      [55]
        bool bMarked
        jointRx jJointRx = {j1=119.753729, j2=-7.953574, j3=74.820625, j4=-173.223401, j5=72.415611, j6=-212.309715}
        pointRx pInter
        paraItem pParaItem
          [0]
            bool bSafePoint
            ifItem iIfItem
              [0]
                bool bANDOR[2]
                num nSigIndex[3]
                num nSigType[3]
                num nValue[3]
            mdesc mMdesc = {leave=0}
            num nActionIndex = 41
            num nDelay = 1
            num nMoveType = 1
            num nPercentage
            num nSigValue
        pointRx pPointRx[2] = {x=-39.963894, y=381.881422, z=1281.672322, rx=1.496816, ry=8.299138, rz=89.69815, shoulder=lefty, elbow=epositive, wrist=wpositive}
        string sID
      [56]
        bool bMarked
        jointRx jJointRx = {j1=126.372801, j2=0.947016, j3=58.247522, j4=-173.633502, j5=65.467797, j6=-219.528921}
        pointRx pInter
        paraItem pParaItem
          [0]
            bool bSafePoint
            ifItem iIfItem
              [0]
                bool bANDOR[2]
                num nSigIndex[3]
                num nSigType[3]
                num nValue[3]
            mdesc mMdesc = {leave=0}
            num nActionIndex = 41
            num nDelay = 1
            num nMoveType = 1
            num nPercentage
            num nSigValue
        pointRx pPointRx[2] = {x=-110.0468221, y=381.881454, z=1352.0109929, rx=1.496598, ry=8.298005, rz=89.698483, shoulder=lefty, elbow=epositive, wrist=wpositive}
        string sID
      [57]
        bool bMarked
        jointRx jJointRx = {j1=135.765404, j2=12.255762, j3=45.397511, j4=-174.78792, j5=64.742909, j6=-228.47546}
        pointRx pInter
        paraItem pParaItem
          [0]
            bool bSafePoint
            ifItem iIfItem
              [0]
                bool bANDOR[2]
                num nSigIndex[3]
                num nSigType[3]
                num nValue[3]
            mdesc mMdesc = {leave=0}
            num nActionIndex = 41
            num nDelay = 1
            num nMoveType = 1
            num nPercentage
            num nSigValue
        pointRx pPointRx[2] = {x=-234.761691, y=381.497821, z=1353.29132, rx=1.49622, ry=8.29735, rz=89.698646, shoulder=lefty, elbow=epositive, wrist=wpositive}
        string sID
      [58]
        bool bMarked
        jointRx jJointRx = {j1=138.772753, j2=12.465275, j3=53.540842, j4=-175.467559, j5=73.29136, j6=-230.546088}
        pointRx pInter
        paraItem pParaItem
          [0]
            bool bSafePoint
            ifItem iIfItem
              [0]
                bool bANDOR[2]
                num nSigIndex[3]
                num nSigType[3]
                num nValue[3]
            mdesc mMdesc = {leave=0}
            num nActionIndex = 41
            num nDelay = 1
            num nMoveType = 1
            num nPercentage
            num nSigValue
        pointRx pPointRx[2] = {x=-284.713057, y=381.881445, z=1282.27146, rx=1.496715, ry=8.298986, rz=89.698256, shoulder=lefty, elbow=epositive, wrist=wpositive}
        string sID
      [59]
        bool bMarked
        jointRx jJointRx = {j1=142.602482, j2=20.481815, j3=43.70957, j4=-175.946983, j5=71.740182, j6=-234.319694}
        pointRx pInter
        paraItem pParaItem
          [0]
            bool bSafePoint
            ifItem iIfItem
              [0]
                bool bANDOR[2]
                num nSigIndex[3]
                num nSigType[3]
                num nValue[3]
            mdesc mMdesc = {leave=0}
            num nActionIndex = 41
            num nDelay = 1
            num nMoveType = 1
            num nPercentage
            num nSigValue
        pointRx pPointRx[2] = {x=-357.530662, y=381.881364, z=1278.257011, rx=1.496095, ry=8.297308, rz=89.698645, shoulder=lefty, elbow=epositive, wrist=wpositive}
        string sID
      [60]
        bool bMarked
        jointRx jJointRx = {j1=146.225971, j2=34.147401, j3=22.485673, j4=-176.265369, j5=64.412135, j6=-238.261186}
        pointRx pInter
        paraItem pParaItem
          [0]
            bool bSafePoint
            ifItem iIfItem
              [0]
                bool bANDOR[2]
                num nSigIndex[3]
                num nSigType[3]
                num nValue[3]
            mdesc mMdesc = {leave=0}
            num nActionIndex = 41
            num nDelay = 1
            num nMoveType = 1
            num nPercentage
            num nSigValue
        pointRx pPointRx[2] = {x=-439.57558, y=381.88118, z=1286.715302, rx=1.495603, ry=8.296388, rz=89.698782, shoulder=lefty, elbow=epositive, wrist=wpositive}
        string sID
      [61]
        bool bMarked
        jointRx jJointRx = {j1=145.163516, j2=25.787023, j3=46.647021, j4=-176.436157, j5=80.123032, j6=-236.204112}
        pointRx pInter
        paraItem pParaItem
          [0]
            bool bSafePoint
            ifItem iIfItem
              [0]
                bool bANDOR[2]
                num nSigIndex[3]
                num nSigType[3]
                num nValue[3]
            mdesc mMdesc = {leave=0}
            num nActionIndex = 41
            num nDelay = 1
            num nMoveType = 1
            num nPercentage
            num nSigValue
        pointRx pPointRx[2] = {x=-433.595736, y=395.563274, z=1186.609873, rx=1.496133, ry=8.298356, rz=89.698378, shoulder=lefty, elbow=epositive, wrist=wpositive}
        string sID
      [62]
        bool bMarked
        jointRx jJointRx = {j1=141.740249, j2=16.896756, j3=58.529423, j4=-176.00804128, j5=82.891986, j6=-232.685997}
        pointRx pInter
        paraItem pParaItem
          [0]
            bool bSafePoint
            ifItem iIfItem
              [0]
                bool bANDOR[2]
                num nSigIndex[3]
                num nSigType[3]
                num nValue[3]
            mdesc mMdesc = {leave=0}
            num nActionIndex = 41
            num nDelay = 1
            num nMoveType = 1
            num nPercentage
            num nSigValue
        pointRx pPointRx[2] = {x=-357.383669, y=395.563229, z=1187.219278, rx=1.496378, ry=8.298339, rz=89.698402, shoulder=lefty, elbow=epositive, wrist=wpositive}
        string sID
      [63]
        bool bMarked
        jointRx jJointRx = {j1=145.520586, j2=24.877498, j3=53.652175, j4=-176.529516, j5=86.228461, j6=-236.175028}
        pointRx pInter
        paraItem pParaItem
          [0]
            bool bSafePoint
            ifItem iIfItem
              [0]
                bool bANDOR[2]
                num nSigIndex[3]
                num nSigType[3]
                num nValue[3]
            mdesc mMdesc = {leave=0}
            num nActionIndex = 41
            num nDelay = 1
            num nMoveType = 1
            num nPercentage
            num nSigValue
        pointRx pPointRx[2] = {x=-442.31911, y=395.563141, z=1133.387458, rx=1.496409, ry=8.298276, rz=89.698428, shoulder=lefty, elbow=epositive, wrist=wpositive}
        string sID
      [64]
        bool bMarked
        jointRx jJointRx = {j1=142.932218, j2=18.224798, j3=62.561776, j4=-176.192349, j5=88.31967, j6=-233.487703}
        pointRx pInter
        paraItem pParaItem
          [0]
            bool bSafePoint
            ifItem iIfItem
              [0]
                bool bANDOR[2]
                num nSigIndex[3]
                num nSigType[3]
                num nValue[3]
            mdesc mMdesc = {leave=0}
            num nActionIndex = 41
            num nDelay = 1
            num nMoveType = 1
            num nPercentage
            num nSigValue
        pointRx pPointRx[2] = {x=-383.080032, y=395.992805, z=1133.387618, rx=1.496541, ry=8.298786, rz=89.698287, shoulder=lefty, elbow=epositive, wrist=wpositive}
        string sID
      [65]
        bool bMarked
        jointRx jJointRx = {j1=137.828285, j2=8.0182986, j3=75.0979146, j4=-175.541144, j5=90.27829, j6=-228.278804}
        pointRx pInter
        paraItem pParaItem
          [0]
            bool bSafePoint
            ifItem iIfItem
              [0]
                bool bANDOR[2]
                num nSigIndex[3]
                num nSigType[3]
                num nValue[3]
            mdesc mMdesc = {leave=0}
            num nActionIndex = 41
            num nDelay = 1
            num nMoveType = 1
            num nPercentage
            num nSigValue
        pointRx pPointRx[2] = {x=-282.0829755, y=394.174282, z=1131.442193, rx=1.496419, ry=8.298256, rz=89.698436, shoulder=lefty, elbow=epositive, wrist=wpositive}
        string sID
      [66]
        bool bMarked
        jointRx jJointRx = {j1=129.569522, j2=-2.763661, j3=86.443161, j4=-174.560173, j5=90.131021, j6=-220.057051}
        pointRx pInter
        paraItem pParaItem
          [0]
            bool bSafePoint
            ifItem iIfItem
              [0]
                bool bANDOR[2]
                num nSigIndex[3]
                num nSigType[3]
                num nValue[3]
            mdesc mMdesc = {leave=0}
            num nActionIndex = 41
            num nDelay = 1
            num nMoveType = 1
            num nPercentage
            num nSigValue
        pointRx pPointRx[2] = {x=-158.339339, y=393.754355, z=1130.374707, rx=1.496575, ry=8.298917, rz=89.698258, shoulder=lefty, elbow=epositive, wrist=wpositive}
        string sID
      [67]
        bool bMarked
        jointRx jJointRx = {j1=127.108283, j2=-4.31187, j3=84.0279326, j4=-174.275111, j5=85.948662, j6=-218.0171002}
        pointRx pInter
        paraItem pParaItem
          [0]
            bool bSafePoint
            ifItem iIfItem
              [0]
                bool bANDOR[2]
                num nSigIndex[3]
                num nSigType[3]
                num nValue[3]
            mdesc mMdesc = {leave=0}
            num nActionIndex = 41
            num nDelay = 1
            num nMoveType = 1
            num nPercentage
            num nSigValue
        pointRx pPointRx[2] = {x=-128.944462, y=395.563233, z=1167.186243, rx=1.496331, ry=8.29773, rz=89.69859, shoulder=lefty, elbow=epositive, wrist=wpositive}
        string sID
      [68]
        bool bMarked
        jointRx jJointRx = {j1=127.132916, j2=-2.202885, j3=74.171846, j4=-174.169676, j5=78.242682, j6=-218.827696}
        pointRx pInter
        paraItem pParaItem
          [0]
            bool bSafePoint
            ifItem iIfItem
              [0]
                bool bANDOR[2]
                num nSigIndex[3]
                num nSigType[3]
                num nValue[3]
            mdesc mMdesc = {leave=0}
            num nActionIndex = 41
            num nDelay = 1
            num nMoveType = 1
            num nPercentage
            num nSigValue
        pointRx pPointRx[2] = {x=-129.246182, y=395.563221, z=1240.287458, rx=1.496095, ry=8.297201, rz=89.698751, shoulder=lefty, elbow=epositive, wrist=wpositive}
        string sID
      [69]
        bool bMarked
        jointRx jJointRx = {j1=119.726319, j2=-8.925081, j3=83.332444, j4=-173.436836, j5=79.901655, j6=-211.381836}
        pointRx pInter
        paraItem pParaItem
          [0]
            bool bSafePoint
            ifItem iIfItem
              [0]
                bool bANDOR[2]
                num nSigIndex[3]
                num nSigType[3]
                num nValue[3]
            mdesc mMdesc = {leave=0}
            num nActionIndex = 41
            num nDelay = 1
            num nMoveType = 1
            num nPercentage
            num nSigValue
        pointRx pPointRx[2] = {x=-47.509267, y=395.563233, z=1212.190941, rx=1.496528, ry=8.298847, rz=89.698245, shoulder=lefty, elbow=epositive, wrist=wpositive}
        string sID
      [70]
        bool bMarked
        jointRx jJointRx = {j1=117.0356638, j2=-11.369619, j3=88.345877, j4=-173.227501, j5=82.15053, j6=-208.458383}
        pointRx pInter
        paraItem pParaItem
          [0]
            bool bSafePoint
            ifItem iIfItem
              [0]
                bool bANDOR[2]
                num nSigIndex[3]
                num nSigType[3]
                num nValue[3]
            mdesc mMdesc = {leave=0}
            num nActionIndex = 41
            num nDelay = 1
            num nMoveType = 1
            num nPercentage
            num nSigValue
        pointRx pPointRx[2] = {x=-21.101146, y=395.563202, z=1184.53881, rx=1.49646, ry=8.299163, rz=89.698163, shoulder=lefty, elbow=epositive, wrist=wpositive}
        string sID
      [71]
        bool bMarked
        jointRx jJointRx = {j1=111.636883, j2=-14.155418, j3=90.562702, j4=-172.749065, j5=80.943983, j6=-203.256882}
        pointRx pInter
        paraItem pParaItem
          [0]
            bool bSafePoint
            ifItem iIfItem
              [0]
                bool bANDOR[2]
                num nSigIndex[3]
                num nSigType[3]
                num nValue[3]
            mdesc mMdesc = {leave=0}
            num nActionIndex = 41
            num nDelay = 1
            num nMoveType = 1
            num nPercentage
            num nSigValue
        pointRx pPointRx[2] = {x=27.98203, y=395.563196, z=1184.484299, rx=1.496405, ry=8.299077, rz=89.698195, shoulder=lefty, elbow=epositive, wrist=wpositive}
        string sID
      [72]
        bool bMarked
        jointRx jJointRx = {j1=102.0811227, j2=-15.748657, j3=85.809651, j4=-171.860362, j5=73.429784, j6=-194.828465}
        pointRx pInter
        paraItem pParaItem
          [0]
            bool bSafePoint
            ifItem iIfItem
              [0]
                bool bANDOR[2]
                num nSigIndex[3]
                num nSigType[3]
                num nValue[3]
            mdesc mMdesc = {leave=0}
            num nActionIndex = 41
            num nDelay = 1
            num nMoveType = 1
            num nPercentage
            num nSigValue
        pointRx pPointRx[2] = {x=105.742398, y=395.563206, z=1239.205231, rx=1.496267, ry=8.297338, rz=89.69876, shoulder=lefty, elbow=epositive, wrist=wpositive}
        string sID
      [73]
        bool bMarked
        jointRx jJointRx = {j1=101.965226, j2=-17.946235, j3=95.328716, j4=-172.0869886, j5=80.664903, j6=-193.668084}
        pointRx pInter
        paraItem pParaItem
          [0]
            bool bSafePoint
            ifItem iIfItem
              [0]
                bool bANDOR[2]
                num nSigIndex[3]
                num nSigType[3]
                num nValue[3]
            mdesc mMdesc = {leave=0}
            num nActionIndex = 41
            num nDelay = 1
            num nMoveType = 1
            num nPercentage
            num nSigValue
        pointRx pPointRx[2] = {x=106.315326, y=397.144334, z=1166.222142, rx=1.496509, ry=8.299055, rz=89.698157, shoulder=lefty, elbow=epositive, wrist=wpositive}
        string sID
      [74]
        bool bMarked
        jointRx jJointRx = {j1=109.159845, j2=-17.523216, j3=103.974266, j4=-172.590397, j5=90.481549, j6=-198.656551}
        pointRx pInter
        paraItem pParaItem
          [0]
            bool bSafePoint
            ifItem iIfItem
              [0]
                bool bANDOR[2]
                num nSigIndex[3]
                num nSigType[3]
                num nValue[3]
            mdesc mMdesc = {leave=0}
            num nActionIndex = 41
            num nDelay = 1
            num nMoveType = 1
            num nPercentage
            num nSigValue
        pointRx pPointRx[2] = {x=50.737737, y=395.235981, z=1081.2527, rx=1.365617, ry=8.320655, rz=90.602673, shoulder=lefty, elbow=epositive, wrist=wpositive}
        string sID
      [75]
        bool bMarked
        jointRx jJointRx = {j1=127.797119, j2=-7.36114, j3=94.145293, j4=-174.260119, j5=92.961428, j6=-217.108293}
        pointRx pInter
        paraItem pParaItem
          [0]
            bool bSafePoint
            ifItem iIfItem
              [0]
                bool bANDOR[2]
                num nSigIndex[3]
                num nSigType[3]
                num nValue[3]
            mdesc mMdesc = {leave=0}
            num nActionIndex = 41
            num nDelay = 1
            num nMoveType = 1
            num nPercentage
            num nSigValue
        pointRx pPointRx[2] = {x=-122.311347, y=380.240336, z=1097.145793, rx=1.366321, ry=8.319807, rz=90.60222, shoulder=lefty, elbow=epositive, wrist=wpositive}
        string sID
      [76]
        bool bMarked
        jointRx jJointRx = {j1=125.779161, j2=-6.385537, j3=105.0494702, j4=-173.853648, j5=104.570742, j6=-213.837709}
        pointRx pInter
        paraItem pParaItem
          [0]
            bool bSafePoint
            ifItem iIfItem
              [0]
                bool bANDOR[2]
                num nSigIndex[3]
                num nSigType[3]
                num nValue[3]
            mdesc mMdesc = {leave=0}
            num nActionIndex = 41
            num nDelay = 1
            num nMoveType = 1
            num nPercentage
            num nSigValue
        pointRx pPointRx[2] = {x=-110.0368459, y=395.408133, z=984.452829, rx=1.365734, ry=8.321441, rz=90.601591, shoulder=lefty, elbow=epositive, wrist=wpositive}
        string sID
      [77]
        bool bMarked
        jointRx jJointRx = {j1=119.326527, j2=-11.582985, j3=109.490487, j4=-173.241478, j5=103.100713, j6=-207.390601}
        pointRx pInter
        paraItem pParaItem
          [0]
            bool bSafePoint
            ifItem iIfItem
              [0]
                bool bANDOR[2]
                num nSigIndex[3]
                num nSigType[3]
                num nValue[3]
            mdesc mMdesc = {leave=0}
            num nActionIndex = 41
            num nDelay = 1
            num nMoveType = 1
            num nPercentage
            num nSigValue
        pointRx pPointRx[2] = {x=-40.591401, y=394.609819, z=984.558922, rx=1.365882, ry=8.32114, rz=90.601792, shoulder=lefty, elbow=epositive, wrist=wpositive}
        string sID
      [78]
        bool bMarked
        jointRx jJointRx = {j1=132.430725, j2=-0.0105859, j3=95.557924, j4=-174.666115, j5=102.128999, j6=-220.90754}
        pointRx pInter
        paraItem pParaItem
          [0]
            bool bSafePoint
            ifItem iIfItem
              [0]
                bool bANDOR[2]
                num nSigIndex[3]
                num nSigType[3]
                num nValue[3]
            mdesc mMdesc = {leave=0}
            num nActionIndex = 41
            num nDelay = 1
            num nMoveType = 1
            num nPercentage
            num nSigValue
        pointRx pPointRx[2] = {x=-194.801487, y=395.23596, z=1017.247506, rx=1.365663, ry=8.319364, rz=90.602406, shoulder=lefty, elbow=epositive, wrist=wpositive}
        string sID
      [79]
        bool bMarked
        jointRx jJointRx = {j1=132.458828, j2=-0.0790471, j3=87.268524, j4=-174.777202, j5=93.809024, j6=-221.71153}
        pointRx pInter
        paraItem pParaItem
          [0]
            bool bSafePoint
            ifItem iIfItem
              [0]
                bool bANDOR[2]
                num nSigIndex[3]
                num nSigType[3]
                num nValue[3]
            mdesc mMdesc = {leave=0}
            num nActionIndex = 41
            num nDelay = 1
            num nMoveType = 1
            num nPercentage
            num nSigValue
        pointRx pPointRx[2] = {x=-195.890159, y=395.991481, z=1097.382802, rx=1.365665, ry=8.319356, rz=90.602356, shoulder=lefty, elbow=epositive, wrist=wpositive}
        string sID
      [80]
        bool bMarked
        jointRx jJointRx = {j1=140.806129, j2=12.0425255, j3=73.960822, j4=-175.797158, j5=93.312882, j6=-230.129694}
        pointRx pInter
        paraItem pParaItem
          [0]
            bool bSafePoint
            ifItem iIfItem
              [0]
                bool bANDOR[2]
                num nSigIndex[3]
                num nSigType[3]
                num nValue[3]
            mdesc mMdesc = {leave=0}
            num nActionIndex = 41
            num nDelay = 1
            num nMoveType = 1
            num nPercentage
            num nSigValue
        pointRx pPointRx[2] = {x=-331.291278, y=393.580774, z=1097.744174, rx=1.365543, ry=8.319675, rz=90.602254, shoulder=lefty, elbow=epositive, wrist=wpositive}
        string sID
      [81]
        bool bMarked
        jointRx jJointRx = {j1=140.705878, j2=12.192026, j3=82.155939, j4=-175.702495, j5=101.628566, j6=-229.405986}
        pointRx pInter
        paraItem pParaItem
          [0]
            bool bSafePoint
            ifItem iIfItem
              [0]
                bool bANDOR[2]
                num nSigIndex[3]
                num nSigType[3]
                num nValue[3]
            mdesc mMdesc = {leave=0}
            num nActionIndex = 41
            num nDelay = 1
            num nMoveType = 1
            num nPercentage
            num nSigValue
        pointRx pPointRx[2] = {x=-331.364201, y=395.235947, z=1017.432775, rx=1.365957, ry=8.321078, rz=90.601815, shoulder=lefty, elbow=epositive, wrist=wpositive}
        string sID
      [82]
        bool bMarked
        jointRx jJointRx = {j1=141.483674, j2=14.580293, j3=86.0660414, j4=-182.560432, j5=99.634816, j6=-231.106968}
        pointRx pInter
        paraItem pParaItem
          [0]
            bool bSafePoint
            ifItem iIfItem
              [0]
                bool bANDOR[2]
                num nSigIndex[3]
                num nSigType[3]
                num nValue[3]
            mdesc mMdesc = {leave=0}
            num nActionIndex = 41
            num nDelay = 1
            num nMoveType = 1
            num nPercentage
            num nSigValue
        pointRx pPointRx[2] = {x=-456.482312, y=395.0927041, z=988.243024, rx=1.352323, ry=-2.355377, rz=90.855398, shoulder=lefty, elbow=epositive, wrist=wpositive}
        string sID
      [83]
        bool bMarked
        jointRx jJointRx = {j1=46.220955, j2=-26.278248, j3=73.480924, j4=-176.710401, j5=48.400229, j6=-56.2638}
        pointRx pInter
        paraItem pParaItem
          [0]
            bool bSafePoint
            ifItem iIfItem
              [0]
                bool bANDOR[2]
                num nSigIndex[3]
                num nSigType[3]
                num nValue[3]
            mdesc mMdesc = {leave=0}
            num nActionIndex = 41
            num nDelay = 1
            num nMoveType = 1
            num nPercentage
            num nSigValue
        pointRx pPointRx[2] = {x=156.67875, y=334.103919, z=1427.956714, rx=2.532212, ry=0.979884, rz=172.14558, shoulder=lefty, elbow=epositive, wrist=wpositive}
        string sID
      [84]
        bool bMarked
        jointRx jJointRx = {j1=-0.746077, j2=38.654193, j3=103.0610419, j4=-179.633028, j5=123.454226, j6=8.386419}
        pointRx pInter
        paraItem pParaItem
          [0]
            bool bSafePoint
            ifItem iIfItem
              [0]
                bool bANDOR[2]
                num nSigIndex[3]
                num nSigType[3]
                num nValue[3]
            mdesc mMdesc = {leave=10}
            num nActionIndex = 41
            num nDelay = 1
            num nMoveType = 1
            num nPercentage
            num nSigValue
        pointRx pPointRx[2] = {x=872.305806, y=193.820048, z=536.464849, rx=0.56853, ry=18.254398, rz=-172.702509, shoulder=lefty, elbow=epositive, wrist=wpositive}
        string sID
      [85]
        bool bMarked
        jointRx jJointRx = {j1=-0.746077, j2=38.654193, j3=103.0610419, j4=-179.633028, j5=123.454226, j6=8.386419}
        pointRx pInter
        paraItem pParaItem
          [0]
            bool bSafePoint
            ifItem iIfItem
              [0]
                bool bANDOR[2]
                num nSigIndex[3]
                num nSigType[3]
                num nValue[3]
            mdesc mMdesc = {leave=10}
            num nActionIndex = 70
            num nDelay = 1
            num nMoveType = 4
            num nPercentage
            num nSigValue
        pointRx pPointRx[2] = {x=872.305806, y=193.820048, z=536.464849, rx=0.56853, ry=18.254398, rz=-172.702509, shoulder=lefty, elbow=epositive, wrist=wpositive}
        string sID
      [86]
        bool bMarked
        jointRx jJointRx = {j1=-0.746077, j2=38.654193, j3=103.0610419, j4=-179.633028, j5=123.454226, j6=8.386419}
        pointRx pInter
        paraItem pParaItem
          [0]
            bool bSafePoint
            ifItem iIfItem
              [0]
                bool bANDOR[2]
                num nSigIndex[3]
                num nSigType[3]
                num nValue[3]
            mdesc mMdesc = {leave=10}
            num nActionIndex = 71
            num nDelay = 1
            num nMoveType = 4
            num nPercentage
            num nSigValue = 1
        pointRx pPointRx[2] = {x=872.305806, y=193.820048, z=536.464849, rx=0.56853, ry=18.254398, rz=-172.702509, shoulder=lefty, elbow=epositive, wrist=wpositive}
        string sID
      [87]
        bool bMarked
        jointRx jJointRx = {j1=-0.746077, j2=38.654193, j3=103.0610419, j4=-179.633028, j5=123.454226, j6=8.386419}
        pointRx pInter
        paraItem pParaItem
          [0]
            bool bSafePoint
            ifItem iIfItem
              [0]
                bool bANDOR[2]
                num nSigIndex[3]
                num nSigType[3]
                num nValue[3]
            mdesc mMdesc = {leave=10}
            num nActionIndex = 71
            num nDelay = 1
            num nMoveType = 3
            num nPercentage
            num nSigValue = 1
        pointRx pPointRx[2] = {x=872.305806, y=193.820048, z=536.464849, rx=0.56853, ry=18.254398, rz=-172.702509, shoulder=lefty, elbow=epositive, wrist=wpositive}
        string sID
      [88]
        bool bMarked
        jointRx jJointRx = {j1=94.696904, j2=-17.194257, j3=77.457422, j4=-178.674473, j5=60.986606, j6=84.00973218}
        pointRx pInter
        paraItem pParaItem
          [0]
            bool bSafePoint
            ifItem iIfItem
              [0]
                bool bANDOR[2]
                num nSigIndex[3]
                num nSigType[3]
                num nValue[3]
            mdesc mMdesc = {leave=0}
            num nActionIndex = 41
            num nDelay = 1
            num nMoveType = 1
            num nPercentage
            num nSigValue
        pointRx pPointRx[2] = {x=-70.0312062, y=207.928659, z=1348.60192, rx=0.619605, ry=1.21397, rz=-0.649688, shoulder=lefty, elbow=epositive, wrist=wpositive}
        string sID
      [89]
        bool bMarked
        jointRx jJointRx = {j1=92.674277, j2=28.288635, j3=29.11318, j4=-178.544553, j5=51.372983, j6=85.586329}
        pointRx pInter
        paraItem pParaItem
          [0]
            bool bSafePoint
            ifItem iIfItem
              [0]
                bool bANDOR[2]
                num nSigIndex[3]
                num nSigType[3]
                num nValue[3]
            mdesc mMdesc = {leave=0}
            num nActionIndex = 41
            num nDelay = 1
            num nMoveType = 1
            num nPercentage
            num nSigValue
        pointRx pPointRx[2] = {x=-78.36515, y=651.672778, z=1350.140243, rx=-6.0840795, ry=0.854567, rz=-0.845265, shoulder=lefty, elbow=epositive, wrist=wpositive}
        string sID
      [90]
        bool bMarked
        jointRx jJointRx = {j1=92.636781, j2=25.765616, j3=38.048827, j4=-178.660828, j5=57.78113, j6=85.818199}
        pointRx pInter
        paraItem pParaItem
          [0]
            bool bSafePoint
            ifItem iIfItem
              [0]
                bool bANDOR[2]
                num nSigIndex[3]
                num nSigType[3]
                num nValue[3]
            mdesc mMdesc = {leave=0}
            num nActionIndex = 41
            num nDelay = 1
            num nMoveType = 1
            num nPercentage
            num nSigValue
        pointRx pPointRx[2] = {x=-78.365129, y=662.319738, z=1306.542009, rx=-6.0858586, ry=0.854378, rz=-0.845299, shoulder=lefty, elbow=epositive, wrist=wpositive}
        string sID
      [91]
        bool bMarked
        jointRx jJointRx = {j1=92.621294, j2=23.968056, j3=44.692986, j4=-178.725951, j5=62.627267, j6=85.961844}
        pointRx pInter
        paraItem pParaItem
          [0]
            bool bSafePoint
            ifItem iIfItem
              [0]
                bool bANDOR[2]
                num nSigIndex[3]
                num nSigType[3]
                num nValue[3]
            mdesc mMdesc = {leave=0}
            num nActionIndex = 41
            num nDelay = 1
            num nMoveType = 1
            num nPercentage
            num nSigValue
        pointRx pPointRx[2] = {x=-78.365131, y=666.835212, z=1270.569018, rx=-6.0847454, ry=0.854504, rz=-0.845277, shoulder=lefty, elbow=epositive, wrist=wpositive}
        string sID
      [92]
        bool bMarked
        jointRx jJointRx = {j1=92.713698, j2=17.804684, j3=59.507036, j4=-178.795122, j5=71.278521, j6=86.0690239}
        pointRx pInter
        paraItem pParaItem
          [0]
            bool bSafePoint
            ifItem iIfItem
              [0]
                bool bANDOR[2]
                num nSigIndex[3]
                num nSigType[3]
                num nValue[3]
            mdesc mMdesc = {leave=0}
            num nActionIndex = 41
            num nDelay = 1
            num nMoveType = 1
            num nPercentage
            num nSigValue
        pointRx pPointRx[2] = {x=-78.365141, y=640.766438, z=1210.403131, rx=-6.0840607, ry=0.854555, rz=-0.845261, shoulder=lefty, elbow=epositive, wrist=wpositive}
        string sID
      [93]
        bool bMarked
        jointRx jJointRx = {j1=96.554748, j2=-20.665236, j3=76.89328, j4=-167.849866, j5=22.269651, j6=72.482149}
        pointRx pInter
        paraItem pParaItem
          [0]
            bool bSafePoint
            ifItem iIfItem
              [0]
                bool bANDOR[2]
                num nSigIndex[3]
                num nSigType[3]
                num nValue[3]
            mdesc mMdesc = {leave=0}
            num nActionIndex = 41
            num nDelay = 1
            num nMoveType = 1
            num nPercentage
            num nSigValue
        pointRx pPointRx[2] = {x=-80.825183, y=532.545303, z=1358.0265888, rx=-34.666311, ry=0.85591, rz=-0.845314, shoulder=lefty, elbow=epositive, wrist=wpositive}
        string sID
      [94]
        bool bMarked
        jointRx jJointRx = {j1=93.634054, j2=-0.200585, j3=81.614575, j4=-178.59677, j5=73.693191, j6=85.159231}
        pointRx pInter
        paraItem pParaItem
          [0]
            bool bSafePoint
            ifItem iIfItem
              [0]
                bool bANDOR[2]
                num nSigIndex[3]
                num nSigType[3]
                num nValue[3]
            mdesc mMdesc = {leave=0}
            num nActionIndex = 41
            num nDelay = 1
            num nMoveType = 1
            num nPercentage
            num nSigValue
        pointRx pPointRx[2] = {x=-80.825264, y=510.591299, z=1198.230863, rx=-7.794676, ry=0.855921, rz=-0.845268, shoulder=lefty, elbow=epositive, wrist=wpositive}
        string sID
      [95]
        bool bMarked
        jointRx jJointRx = {j1=93.787667, j2=-1.0430847, j3=74.536099, j4=-178.500668, j5=65.779142, j6=84.785838}
        pointRx pInter
        paraItem pParaItem
          [0]
            bool bSafePoint
            ifItem iIfItem
              [0]
                bool bANDOR[2]
                num nSigIndex[3]
                num nSigType[3]
                num nValue[3]
            mdesc mMdesc = {leave=0}
            num nActionIndex = 41
            num nDelay = 1
            num nMoveType = 1
            num nPercentage
            num nSigValue
        pointRx pPointRx[2] = {x=-80.825258, y=486.544321, z=1272.31133, rx=-7.794062, ry=0.855867, rz=-0.845241, shoulder=lefty, elbow=epositive, wrist=wpositive}
        string sID
      [96]
        bool bMarked
        jointRx jJointRx = {j1=91.611305, j2=21.697472, j3=62.831671, j4=-180.107091, j5=81.0880083, j6=86.831666}
        pointRx pInter
        paraItem pParaItem
          [0]
            bool bSafePoint
            ifItem iIfItem
              [0]
                bool bANDOR[2]
                num nSigIndex[3]
                num nSigType[3]
                num nValue[3]
            mdesc mMdesc = {leave=0}
            num nActionIndex = 41
            num nDelay = 1
            num nMoveType = 1
            num nPercentage
            num nSigValue
        pointRx pPointRx[2] = {x=-78.500982, y=656.948047, z=1125.500806, rx=-3.436823, ry=-0.20246, rz=-1.576516, shoulder=lefty, elbow=epositive, wrist=wpositive}
        string sID
      [97]
        bool bMarked
        jointRx jJointRx = {j1=91.74229, j2=14.792839, j3=68.296964, j4=-180.0995398, j5=79.648805, j6=86.702226}
        pointRx pInter
        paraItem pParaItem
          [0]
            bool bSafePoint
            ifItem iIfItem
              [0]
                bool bANDOR[2]
                num nSigIndex[3]
                num nSigType[3]
                num nValue[3]
            mdesc mMdesc = {leave=0}
            num nActionIndex = 41
            num nDelay = 1
            num nMoveType = 1
            num nPercentage
            num nSigValue
        pointRx pPointRx[2] = {x=-78.500976, y=598.124362, z=1158.0889668, rx=-3.436454, ry=-0.202433, rz=-1.576501, shoulder=lefty, elbow=epositive, wrist=wpositive}
        string sID
      [98]
        bool bMarked
        jointRx jJointRx = {j1=92.0280436, j2=9.342775, j3=74.786055, j4=-180.0818129, j5=80.688357, j6=86.412375}
        pointRx pInter
        paraItem pParaItem
          [0]
            bool bSafePoint
            ifItem iIfItem
              [0]
                bool bANDOR[2]
                num nSigIndex[3]
                num nSigType[3]
                num nValue[3]
            mdesc mMdesc = {leave=0}
            num nActionIndex = 41
            num nDelay = 1
            num nMoveType = 1
            num nPercentage
            num nSigValue
        pointRx pPointRx[2] = {x=-80.49317, y=552.392448, z=1158.114787, rx=-3.435481, ry=-0.202365, rz=-1.576463, shoulder=lefty, elbow=epositive, wrist=wpositive}
        string sID
      [99]
        bool bMarked
        jointRx jJointRx = {j1=92.249877, j2=2.333444, j3=85.899577, j4=-180.0676659, j5=84.792822, j6=86.183874}
        pointRx pInter
        paraItem pParaItem
          [0]
            bool bSafePoint
            ifItem iIfItem
              [0]
                bool bANDOR[2]
                num nSigIndex[3]
                num nSigType[3]
                num nValue[3]
            mdesc mMdesc = {leave=0}
            num nActionIndex = 41
            num nDelay = 1
            num nMoveType = 1
            num nPercentage
            num nSigValue
        pointRx pPointRx[2] = {x=-80.825194, y=493.950637, z=1125.0300688, rx=-3.434917, ry=-0.202308, rz=-1.576433, shoulder=lefty, elbow=epositive, wrist=wpositive}
        string sID
      [100]
        bool bMarked
        jointRx jJointRx = {j1=92.358026, j2=-0.641957, j3=96.255336, j4=-180.060943, j5=92.172944, j6=86.067457}
        pointRx pInter
        paraItem pParaItem
          [0]
            bool bSafePoint
            ifItem iIfItem
              [0]
                bool bANDOR[2]
                num nSigIndex[3]
                num nSigType[3]
                num nValue[3]
            mdesc mMdesc = {leave=0}
            num nActionIndex = 41
            num nDelay = 1
            num nMoveType = 1
            num nPercentage
            num nSigValue
        pointRx pPointRx[2] = {x=-80.825191, y=465.498955, z=1054.656021, rx=-3.435026, ry=-0.202315, rz=-1.576444, shoulder=lefty, elbow=epositive, wrist=wpositive}
        string sID
      [101]
        bool bMarked
        jointRx jJointRx = {j1=92.380346, j2=-0.232216, j3=102.0680251, j4=-180.0600521, j5=98.398016, j6=86.0384955}
        pointRx pInter
        paraItem pParaItem
          [0]
            bool bSafePoint
            ifItem iIfItem
              [0]
                bool bANDOR[2]
                num nSigIndex[3]
                num nSigType[3]
                num nValue[3]
            mdesc mMdesc = {leave=0}
            num nActionIndex = 41
            num nDelay = 1
            num nMoveType = 1
            num nPercentage
            num nSigValue
        pointRx pPointRx[2] = {x=-80.824957, y=459.966175, z=995.666701, rx=-3.432367, ry=-0.202053, rz=-1.576659, shoulder=lefty, elbow=epositive, wrist=wpositive}
        string sID
      [102]
        bool bMarked
        jointRx jJointRx = {j1=92.64202, j2=26.0515396, j3=70.311343, j4=-178.981022, j5=92.852687, j6=86.568019}
        pointRx pInter
        paraItem pParaItem
          [0]
            bool bSafePoint
            ifItem iIfItem
              [0]
                bool bANDOR[2]
                num nSigIndex[3]
                num nSigType[3]
